Staubli VAL3: trajTemp.pjx

--- trajTemp.pjx ---
Parameters version=s8.15.3Cs9_BS3337 stackSize=5000 millimeterUnit=true
Program file=start.pgx
Program file=stop.pgx
Data file=trajTemp.dtx
Type name=trajItem path=Disk://source/template/trajItem/trajItem.pjx

--- trajTemp.dtx ---
public trajItem tTrajItem{}

--- start.pgx ---
program start()
begin
end

--- stop.pgx ---
program stop()
begin
end
